(* IEC 61131-3 sources: 2026_Projet_YGO_ExcavatriceDragage/CODE_BACKUP/CODE_20260822_IntroductionTestCI/G_CYCLE, 6 files *)

(* ---- E_CycleStep.st ---- *)
(* =======================================================================
   ⚙️ E_CycleStep — Étapes de la machine d'état du cycle automatique
   ───────────────────────────────────────────────────────────────
   🎯 Rôle : Énumération des étapes du cycle automatique de dragage (X0 à X13 + STABILIZING)
   📄 Doc métier : DOC/AF/AF_Partie-04_Mode_SemiAuto_Sequenceur_v2.1.md
   ======================================================================= *)

TYPE E_CycleStep :
(
  X0_PREPARATION      := 0,   (* Début de graphe : à la TRÉMIE, treuils en position HAUTE *)
  X1_HOMING           := 1,   (* Vitesses lentes pour chercher capteur top + référencement *)
  X2_WORK_POS_SELECT  := 2,   (* Sélection cible Trémie/P1/Maintenance + translation validée *)
  X3_OPEN_BUCKET      := 3,   (* Ouverture benne (si déjà ouverte -> passe vite) *)
  X4_DESCEND_OPEN     := 4,   (* Plongée benne ouverte, M1+M2 synchro, Kobold mesure ON *)
  X5_BOTTOM_CONFIRMED := 5,   (* Fond validé (FB_DiveSearch) ; arrêt descente *)
  X6_CLOSE_BUCKET     := 6,   (* Fermeture benne — tolérance « à peu près fermé » *)
  X7_CTRL_ASCENT      := 7,   (* Remontée palier 1 de contrôle *)
  X8_ASCENT_LOADED    := 8,   (* Remontée nominale jusqu'à limite haute *)
  X9_DRAIN_PAUSE      := 9,   (* Égouttage temporisé — temps affiché IHM *)
  X10_TRANSLATE_DUMP  := 10,  (* Translation vers trémie + avertissements IHM *)
  X11_OPEN_DUMP       := 11,  (* Ouverture benne = vidage ; montée possible, descente ouvre *)
  X13_DONE_SYNC       := 13,  (* Fin de cycle, synchronisation finale (R4) + compteur *)
  STABILIZING         := 14   (* État d'attente/stabilisation — pas une erreur *)
);
END_TYPE

(* ---- E_DiveSearchState.st ---- *)
(* =======================================================================
   ⚙️ E_DiveSearchState — Phases internes de recherche du fond Kobold
   ───────────────────────────────────────────────────────────────
   🎯 Rôle : Énumération des phases de détection et recherche du fond
   📄 Doc métier : DOC/AF/AF_Partie-04_Mode_SemiAuto_Sequenceur_v2.1.md
   ======================================================================= *)

TYPE E_DiveSearchState :
(
    WAIT_PRECONDITIONS := 0, (* Attente benne ouverte, positions et Kobold au repos *)
    READY_TO_DESCEND   := 1, (* Prêt à assister une demande de descente *)
    SEARCHING_IMMERSION := 2, (* Descente : attente front 0->1 dans fenêtre eau *)
    SEARCHING_BOTTOM    := 3, (* Immersion validée : attente front 1->0 au fond *)
    BOTTOM_CONFIRMED    := 4, (* Fond validé ; extraction peut être demandée *)
    ERROR_HOLD          := 5  (* Séquence invalide, descente assistée interdite *)
);
END_TYPE

(* ---- E_ExtractionSequenceState.st ---- *)
(* =======================================================================
   ⚙️ E_ExtractionSequenceState — Phases d'extraction assistée
   ───────────────────────────────────────────────────────────────
   🎯 Rôle : Énumération des phases de la séquence d'extraction assistée
   📄 Doc métier : DOC/AF/AF_Partie-04_Mode_SemiAuto_Sequenceur_v2.1.md
   ======================================================================= *)

TYPE E_ExtractionSequenceState :
(
    WAIT_BOTTOM_CONFIRMATION := 0, (* Attente fond Kobold ou attestation opérateur *)
    READY_TO_CLOSE            := 1, (* Prêt à fermer la benne *)
    CLOSING_BUCKET            := 2, (* FB_Bucket ferme M2 seul *)
    CONTROL_ASCENT            := 3, (* M1/M2 synchronisés au palier sans contacteur vitesse *)
    NOMINAL_ASCENT            := 4, (* Montée couplée avec vitesse demandée opérateur *)
    ERROR_HOLD                := 5  (* Défaut extraction, reprise interdite avant reset *)
);
END_TYPE

(* ---- FB_Cycle.st ---- *)
(* =======================================================================
   ⚙️ FB_Cycle — Séquenceur du cycle automatique (Grafcet de dragage)
   ───────────────────────────────────────────────────────────────
   🎯 Rôle : Automate de cycle automatique de dragage (X0 à X13 + STABILIZING)
   🔒 Sécurité : Gating par mode et homme-mort, repli STABILIZING sur défaut
   🔌 Interface : Demandes de mouvements (treuils, translation, benne)
   📄 Doc métier : DOC/AF/AF_Partie-04_Mode_SemiAuto_Sequenceur_v2.1.md
   ======================================================================= *)

FUNCTION_BLOCK PUBLIC FB_Cycle
VAR_INPUT
    // === COMMANDES & AUTORISATIONS ===
    Enable                  : BOOL;         // --> [CMD] Activation generale du sequenceur
    Reset                   : BOOL;         // --> [CMD] Acquittement defaut (front)
    PowerContactorEngaged   : BOOL;         // --> [SAFE] Chaine de securite OK
    Mode                    : E_Mode;       // --> [CMD] Mode arbitre (SEMI_AUTO pour instance cycle)
    CycleMotionPermit       : BOOL;         // --> [CMD] Manche deflecte (non centre)
    DeadmanArmed            : BOOL;         // --> [CMD] Appui homme-mort (fenetre 3 s)
    HeartbeatIhmOk          : BOOL;         // --> [SAFE] IHM<->PLC valide

    // === COMMANDES OPERATEUR ===
    StartCycle              : BOOL;         // --> [CMD] Demande lancement / reprise (IHM)
    AbortCycle              : BOOL;         // --> [CMD] Demande abandon (IHM)

    // === CIBLES ET CONFIGURATION ===
    SelTarget               : INT;          // --> [CFG] Cible selectionnee (1=Tremie, 2=P2, 3=P1, 4=Maintenance)
    SetDepthM               : REAL;         // --> [CFG] Profondeur de consigne (negative)
    SetOffsetM              : REAL;         // --> [CFG] Ecart de fermeture benne cible

    // === FEEDBACKS CAPTEURS & MATERIEL ===
    KoboldContactFond       : BOOL;         // --> [HW] Retour dedie Kobold : TRUE = contact fond
    LimitLegalReached       : BOOL;         // --> [SAFE] Limite legale atteinte (descente interdite)
    LimitLegalDepthM        : REAL;         // --> [CFG] Profondeur legale minimale autorisee
    WinchSyncError          : BOOL;         // --> [SAFE] Desynchronisme bloquant M1/M2
    WinchSyncDeltaM         : REAL;         // --> [HW] Ecart codeurs M1/M2 pour diagnostic
    M1_CablePosM            : REAL;         // --> [HW] Position cable treuil M1 (recalee)
    M2_CablePosM            : REAL;         // --> [HW] Position cable treuil M2 (recalee)
    M1_MeasuredSpeedMps     : REAL;         // --> [HW] Vitesse lineaire mesuree M1 (m/s)
    M2_MeasuredSpeedMps     : REAL;         // --> [HW] Vitesse lineaire mesuree M2 (m/s)
    SpeedMismatchThresholdMps : REAL;       // --> [CFG] Seuil ecart vitesse ; 0 = controle desactive
    SpeedMismatchTimeout    : TIME;         // --> [CFG] Duree de confirmation ; 0 = controle desactive
    CableLimitM1AscentM     : REAL;         // --> [CFG] Limite haute d'exploitation M1

    // === FEEDBACKS TRANSLATION M3 ===
    Translation_At_P1           : BOOL;     // --> [HW] Capteur position P1 (arret travail)
    Translation_At_Tremie       : BOOL;     // --> [HW] Capteur fin de course tremie
    Translation_At_Maintenance : BOOL;     // --> [HW] Capteur fin de course maintenance
    Translation_Busy            : BOOL;     // --> [HW] Mouvement translation en cours
    Translation_Done            : BOOL;     // --> [HW] Cible translation atteinte

    // === FEEDBACKS BENNE ===
    Benne_Busy              : BOOL;         // --> [HW] Mouvement machoires benne en cours
    Benne_Done              : BOOL;         // --> [HW] Mouvement ouverture/fermeture termine
    Benne_IsOpen            : BOOL;         // --> [HW] Benne mecaniquement ouverte memorisee
    Benne_IsClosed          : BOOL;         // --> [HW] Benne mecaniquement fermee memorisee
    Benne_IsRoughlyClosed   : BOOL;         // --> [HW] Benne a peu pres fermee (tolerance matiere)

    // === REFERENCEMENT CODEURS ===
    HomedM1                 : BOOL;         // --> [HW] Codeur M1 reference
    HomedM2                 : BOOL;         // --> [HW] Codeur M2 reference
    TopPositionSensor       : BOOL;         // --> [HW] Capteur position haute (referencement)
    HomingRequest           : BOOL;         // --> [CMD] Demande de referencement (front)
END_VAR
VAR_OUTPUT
    // === ETATS IEC & DEFECTUOSITES ===
    Ready                   : BOOL;         // <-- [STAT] Sequenceur disponible
    Busy                    : BOOL;         // <-- [STAT] Cycle automatique actif
    Done                    : BOOL;         // <-- [STAT] Cycle automatique complete
    Error                   : BOOL;         // <-- [STAT] Defaut cycle
    ErrorId                 : WORD;         // <-- [DIAG] Code erreur bitmask
    SpeedMismatchMps        : REAL;         // <-- [DIAG] Ecart absolu vitesse M1/M2 (m/s)
    SpeedMismatchActive     : BOOL;         // <-- [DIAG] Seuil vitesse depasse sur cycle courant
    SpeedMismatchConfirmed  : BOOL;         // <-- [DIAG] Ecart vitesse confirme pendant timeout

    // === ORDRES ACTIONNEURS (COMMANDES STRUCTUREES) ===
    WinchM1Cmd              : ST_WinchCmdDemand;        // <-- [ACT] Demande treuil M1
    WinchM2Cmd              : ST_WinchCmdDemand;        // <-- [ACT] Demande treuil M2
    TranslationCmd          : ST_TranslationCmdDemand;  // <-- [ACT] Demande translation M3
    BucketCmd               : ST_BucketCmdDemand;       // <-- [ACT] Demande benne

    // === METADONNEES & SYNOPTIQUE ===
    CycleStep               : E_CycleStep;  // <-- [STAT] Etape active du Grafcet
    CycleStateStr           : STRING(80);   // <-- [STAT] Libelle en clair de l'etape
    CycleStepAtError        : E_CycleStep;  // <-- [DIAG] Etape specifique au moment du defaut
END_VAR
VAR_IN_OUT
    // === STRUCTURES PARTAGEES & COMPTEURS ===
    SampleCount             : INT;          // <-> [BUS] Compteur de prelevements (RETAIN)
END_VAR
VAR
    // === DETECTEURS DE FRONTS ===
    ResetEdge               : R_TRIG;       // . [LOC] Detecteur front montant Reset
    StartEdge               : R_TRIG;       // . [LOC] Detecteur front montant StartCycle
    DeadmanArmedEdge        : R_TRIG;       // . [LOC] Detecteur front montant DeadmanArmed (demarrage joystick)
    AbortEdge               : R_TRIG;       // . [LOC] Detecteur front montant AbortCycle
    ErrorEdge               : R_TRIG;       // . [LOC] Detecteur front montant Error

    // === ETATS INTERNES ===
    State                   : E_CycleStep := E_CycleStep.X0_PREPARATION; // . [LOC] Etape courante machine d'etat
    SavedState              : E_CycleStep := E_CycleStep.X0_PREPARATION; // . [LOC] Etape memorisee

    // === MEMORISATIONS & REGISTRES INTERNES ===
    TouchPositionM          : REAL;         // . [LOC] Position M1 memorisee lors du contact fond
    RaiseTargetM            : REAL;         // . [LOC] Profondeur de remontee memorisee
    SelectedWorkTarget      : INT;          // . [LOC] Cible de travail memorisee

    // === TEMPORISATEURS INTERNES ===
    DrainingTimer           : TON;          // . [LOC] Temporisateur de vidage (egouttage)
    StabilizationTimer      : TON;          // . [LOC] Temporisation maximale de remontee lente
    SpeedMismatchTimer      : TON;          // . [LOC] Confirmation temporelle ecart de vitesse
    StepMaxTimer            : TON;          // . [LOC] Tempo max d'etape

    // === CONSTANTES & CONFIGURATIONS INTERNES ===
    CtrlAscentDistM         : REAL := 2.0;      // . [LOC] Distance de remontee lente de controle
    CtrlAscentToleranceM    : REAL := 0.25;     // . [LOC] Ecart maximal admis entre codeurs
    CtrlAscentTimeout       : TIME := T#30s;    // . [LOC] Temps max pour zone de stabilisation
    DrainingTime            : TIME := T#5s;     // . [LOC] Temps d'egouttage par defaut
    StepMaxTimeout          : TIME := T#60s;    // . [LOC] Tempo max d'etape
END_VAR

// === IMPLEMENTATION ===

{region "§1 Gate securite"}
// 🛑 1. GATES DE SÉCURITÉ ET BLOCAGE (R8)
IF NOT Enable OR NOT PowerContactorEngaged THEN
    WinchM1Cmd.StartStop   := FALSE;
    WinchM1Cmd.Direction   := 0;
    WinchM1Cmd.SpeedPct    := 0.0;

    WinchM2Cmd.StartStop   := FALSE;
    WinchM2Cmd.Direction   := 0;
    WinchM2Cmd.SpeedPct    := 0.0;

    TranslationCmd.Start   := FALSE;
    TranslationCmd.Target  := 0;

    BucketCmd.Open         := FALSE;
    BucketCmd.Close        := FALSE;
    BucketCmd.KoboldContactorCmd := FALSE;

    State                := E_CycleStep.X0_PREPARATION;   // retour à la PREMIÈRE étape (R8)
    CycleStep            := E_CycleStep.X0_PREPARATION;
    CycleStateStr        := 'X0 - Désactivé : sécurité absente ou auto désactivé';
    Ready                := FALSE;
    Busy                 := FALSE;
    Done                 := FALSE;
    RETURN;
END_IF;
{endregion}

{region "§2 Preparation surveillance et commandes cycle"}
Ready := TRUE;
ResetEdge(CLK := Reset);
StartEdge(CLK := StartCycle);
DeadmanArmedEdge(CLK := DeadmanArmed);
AbortEdge(CLK := AbortCycle);
ErrorEdge(CLK := Error);

// 🧊 R9 — capture l'étape spécifique AVANT la bascule vers STABILIZING
IF ErrorEdge.Q THEN
    CycleStepAtError := State;
END_IF;

// ⏱️ Surveillance indépendante de la remontée lente
StabilizationTimer(IN := (State = E_CycleStep.X7_CTRL_ASCENT), PT := CtrlAscentTimeout);

// 📏 Comparaison vitesse réelle M1/M2
SpeedMismatchMps := ABS(M1_MeasuredSpeedMps - M2_MeasuredSpeedMps);
SpeedMismatchActive := (State = E_CycleStep.X7_CTRL_ASCENT)
                       AND CycleMotionPermit
                       AND (SpeedMismatchThresholdMps > 0.0)
                       AND (SpeedMismatchTimeout > T#0ms)
                       AND (SpeedMismatchMps > SpeedMismatchThresholdMps);
SpeedMismatchTimer(IN := SpeedMismatchActive, PT := SpeedMismatchTimeout);
SpeedMismatchConfirmed := SpeedMismatchTimer.Q;

// Tempo max d'étape (R5) — lancée SEULEMENT si pilotage joystick actif (pas de défaut au repos)
StepMaxTimer(IN := CycleMotionPermit AND (State <> E_CycleStep.X0_PREPARATION)
                  AND (State <> E_CycleStep.X13_DONE_SYNC)
                  AND (State <> E_CycleStep.STABILIZING),
             PT := StepMaxTimeout);

IF ResetEdge.Q THEN
    Error := FALSE;
    ErrorId := 16#0000;
    SavedState := E_CycleStep.X0_PREPARATION;
    IF State = E_CycleStep.STABILIZING THEN
        State := E_CycleStep.X0_PREPARATION;
    END_IF;
END_IF;

// 💓 Perte IHM : repli mémorisé. La reconnexion seule ne relance jamais le cycle.
IF NOT HeartbeatIhmOk AND State <> E_CycleStep.STABILIZING THEN
    Error := TRUE;
    ErrorId := ErrorId OR 16#0020;
    State := E_CycleStep.STABILIZING;
END_IF;

// Défaut de synchronisme : arrêt sûr et acquittement obligatoire.
IF WinchSyncError AND State <> E_CycleStep.STABILIZING THEN
    Error := TRUE;
    ErrorId := ErrorId OR 16#0002;
    State := E_CycleStep.STABILIZING;
END_IF;

// 🛡️ Écart de vitesse confirmé : arrêt du cycle et STABILIZING.
IF SpeedMismatchConfirmed AND State <> E_CycleStep.STABILIZING THEN
    Error := TRUE;
    ErrorId := ErrorId OR 16#0010;
    State := E_CycleStep.STABILIZING;
END_IF;

// Tempo max d'étape dépassée (blocage probable) → défaut
IF StepMaxTimer.Q AND State <> E_CycleStep.STABILIZING THEN
    Error := TRUE;
    ErrorId := ErrorId OR 16#0040;
    State := E_CycleStep.STABILIZING;
END_IF;

// Gestion de l'Abandon (D3 — pas de Pause)
IF AbortEdge.Q THEN
    State := E_CycleStep.X0_PREPARATION;
END_IF;
{endregion}

{region "§3 Machine etat cycle automatique"}
// 🔁 2. LOGIQUE DU SÉQUENCEUR (Machine d'état) — CASE sur enum unique (R1)
CASE State OF

    E_CycleStep.X0_PREPARATION:
        CycleStep := E_CycleStep.X0_PREPARATION;
        CycleStateStr := 'X0 - Vérification cohérence système';
        WinchM1Cmd.StartStop := FALSE; WinchM1Cmd.Direction := 0; WinchM1Cmd.SpeedPct := 0.0;
        WinchM2Cmd.StartStop := FALSE; WinchM2Cmd.Direction := 0; WinchM2Cmd.SpeedPct := 0.0;
        TranslationCmd.Start := FALSE; TranslationCmd.Target := 0;
        BucketCmd.Open := FALSE; BucketCmd.Close := FALSE; BucketCmd.KoboldContactorCmd := FALSE;
        Busy := FALSE; Done := FALSE;

        // Transition si système sain et réarmé (front reset ou démarrage).
        // 🔫 D2 : démarrage par bouton IHM (StartEdge) OU armement homme-mort joystick
        // (DeadmanArmedEdge) — l'opérateur peut lancer depuis l'IHM ou le joystick.
        // La continuité des mouvements ne dépend que de CycleMotionPermit (manche défléchi).
        IF StartEdge.Q OR DeadmanArmedEdge.Q THEN
            State := E_CycleStep.X1_HOMING;
        END_IF;

    E_CycleStep.X1_HOMING:
        CycleStep := E_CycleStep.X1_HOMING;
        CycleStateStr := 'X1 - Référencement codeurs (vitesses lentes)';
        Busy := TRUE;

        // Vitesses lentes pour chercher capteur top + référencement
        IF NOT HomedM1 OR NOT HomedM2 THEN
            WinchM1Cmd.StartStop := CycleMotionPermit;
            WinchM1Cmd.Direction := 1;   // montée lente vers capteur top
            WinchM1Cmd.SpeedPct := 10.0;
            WinchM2Cmd.StartStop := CycleMotionPermit;
            WinchM2Cmd.Direction := 1;
            WinchM2Cmd.SpeedPct := 10.0;
            IF HomingRequest THEN
                // déclenche le référencement (via FB_Encoder_Homing en aval)
                State := E_CycleStep.X2_WORK_POS_SELECT;
            END_IF;
        ELSE
            // déjà homé → passe vite
            State := E_CycleStep.X2_WORK_POS_SELECT;
        END_IF;

    E_CycleStep.X2_WORK_POS_SELECT:
        CycleStep := E_CycleStep.X2_WORK_POS_SELECT;
        CycleStateStr := 'X2 - Sélection position travail';
        Busy := TRUE;

        // Destinations sélectionnables : Trémie(1), P1(3), Maintenance(4).
        // P2(2) n'est PAS une destination — capteur de passage en petite vitesse (PV).
        // Si aucune cible valide n'est sélectionnée, on ATTEND à X2 (pas de défaut) :
        // l'opérateur choisit la position de travail via l'IHM (SelTarget).
        IF (SelTarget = 1) OR (SelTarget = 3) OR (SelTarget = 4) THEN
            SelectedWorkTarget := SelTarget;
            TranslationCmd.Target := SelTarget;
            TranslationCmd.Start := CycleMotionPermit;
            // Arrivée à la cible (Trémie/P1/Maintenance) — capteurs PV/PVP2/P2 = ralentissement
            IF CycleMotionPermit AND (
                (SelTarget = 1 AND Translation_At_Tremie) OR
                (SelTarget = 3 AND Translation_At_P1) OR
                (SelTarget = 4 AND Translation_At_Maintenance)) THEN
                TranslationCmd.Start := FALSE;
                State := E_CycleStep.X3_OPEN_BUCKET;
            END_IF;
        END_IF;

    E_CycleStep.X3_OPEN_BUCKET:
        CycleStep := E_CycleStep.X3_OPEN_BUCKET;
        CycleStateStr := 'X3 - Ouverture benne';
        Busy := TRUE;

        // Ouverture benne ; si déjà ouverte → passe vite
        IF Benne_IsOpen THEN
            State := E_CycleStep.X4_DESCEND_OPEN;
        ELSE
            BucketCmd.Open := CycleMotionPermit;
            IF CycleMotionPermit AND Benne_Done AND Benne_IsOpen THEN
                BucketCmd.Open := FALSE;
                State := E_CycleStep.X4_DESCEND_OPEN;
            END_IF;
        END_IF;

    E_CycleStep.X4_DESCEND_OPEN:
        CycleStep := E_CycleStep.X4_DESCEND_OPEN;
        CycleStateStr := 'X4 - Plongée benne ouverte (synchro)';

        // M1 et M2 descendent ensemble (synchro gérée en aval)
        WinchM1Cmd.StartStop := CycleMotionPermit;
        WinchM1Cmd.Direction := -1;
        WinchM1Cmd.SpeedPct  := 50.0;
        WinchM2Cmd.StartStop := CycleMotionPermit;
        WinchM2Cmd.Direction := -1;
        WinchM2Cmd.SpeedPct  := 50.0;
        BucketCmd.KoboldContactorCmd := TRUE;

        // Transition uniquement sur le retour dédié Kobold.
        IF CycleMotionPermit AND KoboldContactFond THEN
            WinchM1Cmd.StartStop := FALSE;
            WinchM2Cmd.StartStop := FALSE;
            BucketCmd.KoboldContactorCmd := FALSE;
            TouchPositionM := M1_CablePosM;
            IF LimitLegalDepthM < -0.01 THEN
                RaiseTargetM := MAX(TouchPositionM + 0.5, LimitLegalDepthM + 0.5);
            ELSE
                RaiseTargetM := TouchPositionM + 0.5;
            END_IF;
            State := E_CycleStep.X5_BOTTOM_CONFIRMED;
        ELSIF LimitLegalReached THEN
            Error := TRUE;
            ErrorId := ErrorId OR 16#0001;
            WinchM1Cmd.StartStop := FALSE;
            WinchM2Cmd.StartStop := FALSE;
            BucketCmd.KoboldContactorCmd := FALSE;
            State := E_CycleStep.STABILIZING;
        END_IF;

    E_CycleStep.X5_BOTTOM_CONFIRMED:
        CycleStep := E_CycleStep.X5_BOTTOM_CONFIRMED;
        CycleStateStr := 'X5 - Fond confirmé : remontée sécurisée';

        WinchM1Cmd.StartStop := CycleMotionPermit;
        WinchM1Cmd.Direction := 1;
        WinchM1Cmd.SpeedPct := 20.0;
        WinchM2Cmd.StartStop := CycleMotionPermit;
        WinchM2Cmd.Direction := 1;
        WinchM2Cmd.SpeedPct := 20.0;

        // Les deux treuils restent synchronisés jusqu'au-dessus de la limite légale.
        IF CycleMotionPermit AND (M1_CablePosM >= RaiseTargetM) AND (M2_CablePosM >= RaiseTargetM) THEN
            WinchM1Cmd.StartStop := FALSE;
            WinchM2Cmd.StartStop := FALSE;
            State := E_CycleStep.X6_CLOSE_BUCKET;
        END_IF;

    E_CycleStep.X6_CLOSE_BUCKET:
        CycleStep := E_CycleStep.X6_CLOSE_BUCKET;
        CycleStateStr := 'X6 - Fermeture benne (tolérance à peu près fermé)';

        WinchM1Cmd.StartStop := FALSE;
        BucketCmd.Close := TRUE;

        // Tolérance : si benne « à peu près fermée » (matière/objet), on remonte et on contrôle
        IF CycleMotionPermit AND (Benne_Done AND (Benne_IsClosed OR Benne_IsRoughlyClosed)) THEN
            BucketCmd.Close := FALSE;
            State := E_CycleStep.X7_CTRL_ASCENT;
        END_IF;

    E_CycleStep.X7_CTRL_ASCENT:
        CycleStep := E_CycleStep.X7_CTRL_ASCENT;
        CycleStateStr := 'X7 - Remontée lente de contrôle';

        WinchM1Cmd.StartStop := CycleMotionPermit;
        WinchM1Cmd.Direction := 1;
        WinchM1Cmd.SpeedPct  := 20.0;
        WinchM2Cmd.StartStop := CycleMotionPermit;
        WinchM2Cmd.Direction := 1;
        WinchM2Cmd.SpeedPct  := 20.0;

        // Contrôle des deux codeurs
        IF WinchSyncError OR (ABS(M1_CablePosM - M2_CablePosM) > CtrlAscentToleranceM) THEN
            Error := TRUE;
            ErrorId := ErrorId OR 16#0008;
            State := E_CycleStep.STABILIZING;
        ELSIF CycleMotionPermit
           AND (M1_CablePosM >= (TouchPositionM + CtrlAscentDistM))
           AND (M2_CablePosM >= (TouchPositionM + CtrlAscentDistM))
           AND (ABS(M1_CablePosM - M2_CablePosM) <= CtrlAscentToleranceM) THEN
            State := E_CycleStep.X8_ASCENT_LOADED;
        ELSIF StabilizationTimer.Q THEN
            Error := TRUE;
            ErrorId := ErrorId OR 16#0008;
            State := E_CycleStep.STABILIZING;
        END_IF;

    E_CycleStep.X8_ASCENT_LOADED:
        CycleStep := E_CycleStep.X8_ASCENT_LOADED;
        CycleStateStr := 'X8 - Remontée en charge';

        WinchM1Cmd.StartStop := CycleMotionPermit;
        WinchM1Cmd.Direction := 1;
        WinchM1Cmd.SpeedPct  := 70.0;
        WinchM2Cmd.StartStop := CycleMotionPermit;
        WinchM2Cmd.Direction := 1;
        WinchM2Cmd.SpeedPct  := 70.0;

        // Transition alignée sur la limite haute d'exploitation
        IF CycleMotionPermit AND M1_CablePosM >= CableLimitM1AscentM THEN
            WinchM1Cmd.StartStop := FALSE;
            WinchM2Cmd.StartStop := FALSE;
            State := E_CycleStep.X9_DRAIN_PAUSE;
        END_IF;

    E_CycleStep.X9_DRAIN_PAUSE:
        CycleStep := E_CycleStep.X9_DRAIN_PAUSE;
        CycleStateStr := 'X9 - Égouttage du godet en cours';
        WinchM1Cmd.StartStop := FALSE;
        WinchM2Cmd.StartStop := FALSE;

        DrainingTimer(IN := TRUE, PT := DrainingTime);
        // Temps écoulé affiché IHM (CycleStateStr + champ dédié)
        IF CycleMotionPermit AND DrainingTimer.Q THEN
            DrainingTimer(IN := FALSE);
            State := E_CycleStep.X10_TRANSLATE_DUMP;
        END_IF;

    E_CycleStep.X10_TRANSLATE_DUMP:
        CycleStep := E_CycleStep.X10_TRANSLATE_DUMP;
        CycleStateStr := 'X10 - Déplacement vers trémie (grille/crible libres)';

        TranslationCmd.Target := 1; // Trémie
        TranslationCmd.Start := CycleMotionPermit;

        // Avertissement IHM : grille abaissée/libre, crible libre pour réceptionner la charge
        // (porté par CycleStateStr + OperatorAction côté supervision)

        // Transition si translation arrivé à la trémie
        IF CycleMotionPermit AND Translation_At_Tremie THEN
            TranslationCmd.Start := FALSE;
            State := E_CycleStep.X11_OPEN_DUMP;
        END_IF;

    E_CycleStep.X11_OPEN_DUMP:
        CycleStep := E_CycleStep.X11_OPEN_DUMP;
        CycleStateStr := 'X11 - Vidange / ouverture du godet (montée possible, descente ouvre)';

        // Montée possible (treuils vers le haut) ; descente fait ouvrir la benne.
        // Montée : on laisse l'opérateur remonter les 2 treuils en synchro si besoin.
        WinchM1Cmd.StartStop := CycleMotionPermit AND (WinchM1Cmd.Direction = 1);
        WinchM1Cmd.Direction := 1;
        WinchM1Cmd.SpeedPct  := 20.0;
        WinchM2Cmd.StartStop := CycleMotionPermit AND (WinchM2Cmd.Direction = 1);
        WinchM2Cmd.Direction := 1;
        WinchM2Cmd.SpeedPct  := 20.0;

        // Descente → ouverture benne (vidage)
        BucketCmd.Open := CycleMotionPermit AND (WinchM1Cmd.Direction = -1);

        // Contrôle convoyeurs par MESSAGE utilisateur (pas encore câblé) :
        // CycleStateStr + OperatorAction côté supervision demandent de vérifier
        // que les convoyeurs sont en route avant/au lâcher.
        IF CycleMotionPermit AND Benne_Done AND Benne_IsOpen THEN
            BucketCmd.Open := FALSE;
            State := E_CycleStep.X13_DONE_SYNC;
        END_IF;

    E_CycleStep.X13_DONE_SYNC:
        CycleStep := E_CycleStep.X13_DONE_SYNC;
        CycleStateStr := 'X13 - Cycle automatique complété - prêt';
        WinchM1Cmd.StartStop := FALSE;
        WinchM2Cmd.StartStop := FALSE;
        TranslationCmd.Start := FALSE;
        Done := TRUE;
        Busy := FALSE;

        // Compteur de prélèvements (RETAIN, Q3bis) — compte inconditionnellement
        SampleCount := SampleCount + 1;

        // Rebouclage sur X0_PREPARATION (trémie, treuils hauts) — pas de retour P1
        IF StartEdge.Q THEN
            Done := FALSE;
            State := E_CycleStep.X0_PREPARATION;
        END_IF;

    E_CycleStep.STABILIZING:
        CycleStep := E_CycleStep.STABILIZING;
        CycleStateStr := 'X14 - Cycle en attente / stabilisation (STAB)';
        WinchM1Cmd.StartStop := FALSE;
        WinchM2Cmd.StartStop := FALSE;
        TranslationCmd.Start := FALSE;
        BucketCmd.Open := FALSE;
        BucketCmd.Close := FALSE;

END_CASE;
{endregion}

{region "§4 Repli homme mort"}
// 🛑 Relâchement du manche (retour au centre) : aucune demande d'actionneur ne reste active.
// L'étape est mémorisée et reprend au prochain appui valide (D2).
IF Busy AND NOT CycleMotionPermit THEN
    WinchM1Cmd.StartStop := FALSE;
    WinchM2Cmd.StartStop := FALSE;
    TranslationCmd.Start := FALSE;
    BucketCmd.Open := FALSE;
    BucketCmd.Close := FALSE;
    BucketCmd.KoboldContactorCmd := FALSE;
END_IF;
{endregion}

END_FUNCTION_BLOCK

(* ---- FB_DiveSearch.st ---- *)
(* =======================================================================
   ⚙️ FB_DiveSearch — Assistance plongée et recherche du fond Kobold
   ───────────────────────────────────────────────────────────────
   🎯 Rôle : Qualification du capteur Kobold et autorisation de descente
   🛡️ Sécurité : Verrouillage si séquence d'immersion 0->1->0 invalide
   🔌 Interface : Intention de descente et mesures vers permis de descente
   📄 Doc métier : DOC/AF/AF_Partie-04_Mode_SemiAuto_Sequenceur_v2.1.md
   ======================================================================= *)
FUNCTION_BLOCK FB_DiveSearch
VAR_INPUT
    // === COMMANDES & AUTORISATIONS ===
    Enable                  : BOOL;         // --> [CMD] Activation generale du FB (TRUE=Autorise)
    Reset                   : BOOL;         // --> [CMD] Acquittement defaut (front)
    PowerContactorEngaged   : BOOL;         // --> [SAFE] Chaine de securite OK
    Mode                    : E_Mode;       // --> [CMD] Mode de fonctionnement arbitre
    MotionRequestActive     : BOOL;         // --> [CMD] Intention de mouvement active
    MotionDirection         : INT;          // --> [CMD] Sens de mouvement (-1 = descente)

    // === CAPTEURS & ETATS BENNE ===
    BucketIsOpen            : BOOL;         // --> [HW] Benne ouverte confirmee
    KoboldImmersed          : BOOL;         // --> [HW] Capteur Kobold immerge (FALSE=hors eau, TRUE=immerge)
    M1Position_M            : REAL;         // --> [HW] Position codeur treuil M1 (m)
    M2Position_M            : REAL;         // --> [HW] Position codeur treuil M2 (m)
    PositionsValid          : BOOL;         // --> [HW] Validite des mesures de position

    // === CONFIGURATION & SEUILS ===
    DiveStartMin_M          : REAL;         // --> [CFG] Seuil position min pour debut plongee (m)
    ImmersionUpper_M        : REAL;         // --> [CFG] Borne haute fenetre d'immersion (m)
    ImmersionLower_M        : REAL;         // --> [CFG] Borne basse fenetre d'immersion (m)
    BypassPreconditions     : BOOL := FALSE;// --> [TST] Bypass preconditions et seuils (mode test)
END_VAR
VAR_OUTPUT
    // === ETATS IEC & DEFECTUOSITES ===
    Ready                   : BOOL;         // <-- [STAT] FB pret a fonctionner
    // Status.ErrorId : bit0 precond, bit1 seq, bit2 cfg
    Status                  : ST_FbStatus;  // <-- [STAT] Etat global FB (Busy/Done/Error/ErrorId/State/StateAtError)
    DiveState               : E_DiveSearchState; // <-- [STAT] Phase interne de recherche fond

    // === PERMIS & AUTORISATIONS ===
    DescendPermit           : BOOL;         // <-- [ACT] Autorisation de descente assistee
    KoboldMeasureEnable     : BOOL;         // <-- [ACT] Activation mesure/acquisition Kobold
    BottomTouchConfirmed    : BOOL;         // <-- [STAT] Contact fond valide et confirme

    // === DIAGNOSTIC IHM ===
    OperatorActionId        : WORD;         // <-- [DIAG] ID action operateur requise
    OperatorAction          : STRING(120);  // <-- [DIAG] Message explicatif operateur
END_VAR
VAR
    // === DETECTEURS DE FRONTS ===
    ResetEdge               : R_TRIG;       // . [LOC] Detecteur front montant Reset
    KoboldRiseEdge          : R_TRIG;       // . [LOC] Detecteur front entrant eau (0->1)
    KoboldFallEdge          : F_TRIG;       // . [LOC] Detecteur front sortie eau / fond (1->0)

    // === VARIABLES LOCALES INTERNES ===
    ImmersionConfirmed      : BOOL;         // . [LOC] Immersion dans la fenetre d'eau validee
    ErrorCausePresent       : BOOL;         // . [LOC] Presence d'une cause de defaut parametrage
END_VAR

{region "§1 Gate desactivation"}
IF NOT Enable OR NOT PowerContactorEngaged THEN
    Ready := FALSE; Status.Busy := FALSE; Status.Done := FALSE;
    DescendPermit := FALSE; KoboldMeasureEnable := FALSE;
    BottomTouchConfirmed := FALSE;
    Status.State := E_State.DISABLED;
    Status.StateAtError := E_State.DISABLED;
    DiveState := E_DiveSearchState.WAIT_PRECONDITIONS;
    OperatorActionId := 0; OperatorAction := '';
    ImmersionConfirmed := FALSE;
    RETURN;
END_IF;

{endregion}

{region "§2 Preconditions fronts et rearmement"}
ResetEdge(CLK := Reset);
KoboldRiseEdge(CLK := KoboldImmersed);
KoboldFallEdge(CLK := KoboldImmersed);

ErrorCausePresent := NOT BypassPreconditions AND ((DiveStartMin_M < ImmersionUpper_M)
                  OR (ImmersionUpper_M <= ImmersionLower_M));
IF ErrorCausePresent THEN
    Status.ErrorId := Status.ErrorId OR 16#0004;
END_IF;

(* Reset = front + causes disparues ; aucun redémarrage automatique. *)
IF ResetEdge.Q AND NOT ErrorCausePresent AND NOT KoboldImmersed AND NOT MotionRequestActive THEN
    Status.ErrorId := 16#0000;
    ImmersionConfirmed := FALSE;
    BottomTouchConfirmed := FALSE;
    Status.StateAtError := E_State.DISABLED;
    DiveState := E_DiveSearchState.WAIT_PRECONDITIONS;
END_IF;

DescendPermit := FALSE; KoboldMeasureEnable := FALSE;
Ready := FALSE; Status.Busy := FALSE; Status.Done := FALSE;
OperatorActionId := 0; OperatorAction := '';

{endregion}

{region "§3 Machine etat plongee recherche fond"}
IF Status.ErrorId <> 16#0000 THEN
    Status.State := E_State.READY;
    DiveState := E_DiveSearchState.ERROR_HOLD;
    OperatorActionId := 16#0180;
    OperatorAction := 'Vérifier les conditions puis réarmer avant une nouvelle plongée.';
ELSE
    CASE DiveState OF
        E_DiveSearchState.WAIT_PRECONDITIONS:
            Status.State := E_State.INIT;
            IF NOT BypassPreconditions
               AND (NOT BucketIsOpen OR NOT PositionsValid OR KoboldImmersed
                    OR (M1Position_M < DiveStartMin_M) OR (M2Position_M < DiveStartMin_M)) THEN
                OperatorActionId := 16#0100;
                OperatorAction := 'Vérifier les conditions initiales de plongée.';
            ELSE
                DiveState := E_DiveSearchState.READY_TO_DESCEND;
            END_IF;

        E_DiveSearchState.READY_TO_DESCEND:
            Status.State := E_State.READY;
            Ready := TRUE;
            OperatorActionId := 16#0101;
            OperatorAction := 'Demander une descente pour rechercher le fond.';
            IF MotionRequestActive AND (MotionDirection = -1) THEN
                DiveState := E_DiveSearchState.SEARCHING_IMMERSION;
            END_IF;

        E_DiveSearchState.SEARCHING_IMMERSION:
            Status.State := E_State.BUSY;
            Status.Busy := TRUE;
            DescendPermit := MotionRequestActive AND (MotionDirection = -1);
            KoboldMeasureEnable := TRUE;
            OperatorActionId := 16#0102;
            OperatorAction := 'Maintenir la descente : recherche immersion Kobold.';
            IF KoboldRiseEdge.Q THEN
                IF (M1Position_M <= ImmersionUpper_M) AND (M1Position_M >= ImmersionLower_M)
                   AND (M2Position_M <= ImmersionUpper_M) AND (M2Position_M >= ImmersionLower_M) THEN
                    ImmersionConfirmed := TRUE;
                    DiveState := E_DiveSearchState.SEARCHING_BOTTOM;
                ELSE
                    Status.ErrorId := Status.ErrorId OR 16#0002;
                    Status.StateAtError := Status.State;
                END_IF;
            ELSIF (M1Position_M < ImmersionLower_M) OR (M2Position_M < ImmersionLower_M) THEN
                Status.ErrorId := Status.ErrorId OR 16#0002;
                Status.StateAtError := Status.State;
            END_IF;

        E_DiveSearchState.SEARCHING_BOTTOM:
            Status.State := E_State.BUSY;
            Status.Busy := TRUE;
            DescendPermit := MotionRequestActive AND (MotionDirection = -1);
            KoboldMeasureEnable := TRUE;
            OperatorActionId := 16#0103;
            OperatorAction := 'Maintenir la descente : immersion validée, recherche du fond.';
            IF KoboldFallEdge.Q AND ImmersionConfirmed THEN
                BottomTouchConfirmed := TRUE;
                ImmersionConfirmed := FALSE;
                DiveState := E_DiveSearchState.BOTTOM_CONFIRMED;
            END_IF;

        E_DiveSearchState.BOTTOM_CONFIRMED:
            Status.State := E_State.DONE;
            Status.Done := TRUE;
            OperatorActionId := 16#0104;
            OperatorAction := 'Fond détecté : demander la fermeture ou l extraction.';

        E_DiveSearchState.ERROR_HOLD:
            Status.State := E_State.READY;
    END_CASE;
END_IF;

Status.Error := (Status.ErrorId <> 16#0000);

{endregion}

(* ---- FB_ExtractionSequence.st ---- *)
(* =======================================================================
   ⚙️ FB_ExtractionSequence — Fermeture benne et remontée assistée
   ───────────────────────────────────────────────────────────────
   🎯 Rôle : Séquence d'extraction (fermeture benne, remontée de contrôle, remontée nominale)
   🛡️ Sécurité : Aucune remontée assistée sans fond confirmé, contrôle palier 1
   📄 Doc métier : DOC/AF/AF_Partie-04_Mode_SemiAuto_Sequenceur_v2.1.md
   ======================================================================= *)
FUNCTION_BLOCK FB_ExtractionSequence
VAR_INPUT
    // === COMMANDES & AUTORISATIONS ===
    Enable                      : BOOL;     // --> [CMD] Activation generale du FB (TRUE=Autorise)
    Reset                       : BOOL;     // --> [CMD] Acquittement defaut (front)
    PowerContactorEngaged       : BOOL;     // --> [SAFE] Chaine de securite OK
    Mode                        : E_Mode;   // --> [CMD] Mode de fonctionnement arbitre
    MotionRequestActive         : BOOL;     // --> [CMD] Intention de mouvement active
    MotionDirection             : INT;      // --> [CMD] Sens de mouvement (+1 = montee)
    BottomPositionConfirmed     : BOOL;     // --> [SAFE] Attestation fond confirme (Kobold ou op)

    // === CAPTEURS & ETATS MATERIELS ===
    BucketIsClosed              : BOOL;     // --> [HW] Benne fermee confirmee
    BucketBusy                  : BOOL;     // --> [HW] Mouvement benne en cours
    BucketError                 : BOOL;     // --> [SAFE] Defaut sur sous-systeme benne
    WinchSyncError              : BOOL;     // --> [SAFE] Defaut de desynchronisme treuils M1/M2
    M1Position_M                : REAL;     // --> [HW] Position codeur treuil M1 (m)
    M2Position_M                : REAL;     // --> [HW] Position codeur treuil M2 (m)
    M1MeasuredSpeedValid        : BOOL;     // --> [HW] Validite mesure vitesse M1
    M2MeasuredSpeedValid        : BOOL;     // --> [HW] Validite mesure vitesse M2
    PositionsValid              : BOOL;     // --> [HW] Validite des mesures de position

    // === CONFIGURATION & REGLAGES ===
    ControlAscentDistance_M     : REAL;     // --> [CFG] Distance palier 1 de controle remontee (m)
END_VAR
VAR_OUTPUT
    // === ETATS IEC & DEFECTUOSITES ===
    Ready                       : BOOL;     // <-- [STAT] FB pret a fonctionner (sortie libre, hors ST_FbStatus)
    // 🧩 Statut transverse (forme cible) — regroupe Busy/Done/Error/ErrorId/State/StateAtError.
    // ErrorId bit0:fond ; bit1:ferme ; bit2:ctrl ; bit3:cfg.
    Status                      : ST_FbStatus; // <-- [STAT] Etat global FB (Busy/Done/Error/ErrorId/State/StateAtError)
    ExtractionState             : E_ExtractionSequenceState; // <-- [STAT] Phase interne extraction

    // === ORDRES & AUTORISATIONS ===
    BucketCloseRequest          : BOOL;     // <-- [ACT] Demande de fermeture benne
    AscentPermit                : BOOL;     // <-- [ACT] Autorisation de remontee assistee
    ForceMinSpeedStep           : BOOL;     // <-- [ACT] Forcage vitesse minimale (palier de controle)
    BottomConfirmationConsumed  : BOOL;     // <-- [STAT] Signal confirmation fond consomme

    // === DIAGNOSTIC IHM ===
    OperatorActionId            : WORD;     // <-- [DIAG] ID action operateur requise
    OperatorAction              : STRING(120); // <-- [DIAG] Message explicatif operateur
END_VAR
VAR
    // === DETECTEURS DE FRONTS ===
    ResetEdge                   : R_TRIG;   // . [LOC] Detecteur front montant Reset

    // === MEMORISATIONS & POSITIONS INTERNES ===
    ControlStartM1Position_M    : REAL;     // . [LOC] Position M1 au debut du palier de controle (m)
    ControlStartM2Position_M    : REAL;     // . [LOC] Position M2 au debut du palier de controle (m)

    // === VARIABLES LOCALES INTERNES ===
    ErrorCausePresent           : BOOL;     // . [LOC] Presence d'une cause de defaut parametrage
END_VAR

{region "§1 Gate desactivation"}
IF NOT Enable OR NOT PowerContactorEngaged THEN
    Ready := FALSE; Status.Busy := FALSE; Status.Done := FALSE;
    BucketCloseRequest := FALSE; AscentPermit := FALSE; ForceMinSpeedStep := FALSE;
    BottomConfirmationConsumed := FALSE;
    Status.State := E_State.DISABLED;
    Status.StateAtError := E_State.DISABLED;
    ExtractionState := E_ExtractionSequenceState.WAIT_BOTTOM_CONFIRMATION;
    OperatorActionId := 0; OperatorAction := '';
    RETURN;
END_IF;

{endregion}

{region "§2 Preconditions reset et initialisation sorties"}
ResetEdge(CLK := Reset);
ErrorCausePresent := (ControlAscentDistance_M <= 0.0);
IF ErrorCausePresent THEN
    Status.ErrorId := Status.ErrorId OR 16#0008;
END_IF;
IF ResetEdge.Q AND NOT ErrorCausePresent AND NOT MotionRequestActive THEN
    Status.ErrorId := 16#0000;
    Status.StateAtError := E_State.DISABLED;
    ExtractionState := E_ExtractionSequenceState.WAIT_BOTTOM_CONFIRMATION;
END_IF;

Ready := FALSE; Status.Busy := FALSE; Status.Done := FALSE;
BucketCloseRequest := FALSE; AscentPermit := FALSE; ForceMinSpeedStep := FALSE;
BottomConfirmationConsumed := FALSE;
OperatorActionId := 0; OperatorAction := '';

{endregion}

{region "§3 Machine etat fermeture remontee"}
IF Status.ErrorId <> 16#0000 THEN
    Status.State := E_State.READY;
    ExtractionState := E_ExtractionSequenceState.ERROR_HOLD;
    OperatorActionId := 16#0280;
    OperatorAction := 'Vérifier la benne et les treuils puis réarmer avant de reprendre.';
ELSE
    CASE ExtractionState OF
        E_ExtractionSequenceState.WAIT_BOTTOM_CONFIRMATION:
            Status.State := E_State.INIT;
            IF BottomPositionConfirmed THEN
                ExtractionState := E_ExtractionSequenceState.READY_TO_CLOSE;
            ELSE
                OperatorActionId := 16#0200;
                OperatorAction := 'Confirmer que la benne est posée au fond avant extraction.';
            END_IF;

        E_ExtractionSequenceState.READY_TO_CLOSE:
            Status.State := E_State.READY;
            Ready := TRUE;
            OperatorActionId := 16#0201;
            OperatorAction := 'Demander la montée pour fermer la benne.';
            IF MotionRequestActive AND (MotionDirection = 1) THEN
                BottomConfirmationConsumed := TRUE;
                ExtractionState := E_ExtractionSequenceState.CLOSING_BUCKET;
            END_IF;

        E_ExtractionSequenceState.CLOSING_BUCKET:
            Status.State := E_State.BUSY;
            Status.Busy := TRUE;
            BucketCloseRequest := MotionRequestActive AND (MotionDirection = 1);
            OperatorActionId := 16#0202;
            OperatorAction := 'Maintenir la montée : fermeture de la benne en cours.';
            IF BucketError THEN
                Status.ErrorId := Status.ErrorId OR 16#0002;
                Status.StateAtError := Status.State;
            ELSIF BucketIsClosed AND NOT BucketBusy THEN
                ControlStartM1Position_M := M1Position_M;
                ControlStartM2Position_M := M2Position_M;
                ExtractionState := E_ExtractionSequenceState.CONTROL_ASCENT;
            END_IF;

        E_ExtractionSequenceState.CONTROL_ASCENT:
            Status.State := E_State.BUSY;
            Status.Busy := TRUE;
            AscentPermit := MotionRequestActive AND (MotionDirection = 1);
            ForceMinSpeedStep := TRUE;
            OperatorActionId := 16#0203;
            OperatorAction := 'Maintenir la montée : contrôle charge au palier minimal.';
            IF WinchSyncError OR NOT PositionsValid OR NOT M1MeasuredSpeedValid OR NOT M2MeasuredSpeedValid THEN
                Status.ErrorId := Status.ErrorId OR 16#0004;
                Status.StateAtError := Status.State;
            ELSIF (M1Position_M >= (ControlStartM1Position_M + ControlAscentDistance_M))
               AND (M2Position_M >= (ControlStartM2Position_M + ControlAscentDistance_M)) THEN
                ExtractionState := E_ExtractionSequenceState.NOMINAL_ASCENT;
            END_IF;

        E_ExtractionSequenceState.NOMINAL_ASCENT:
            Status.State := E_State.BUSY;
            Status.Busy := TRUE;
            AscentPermit := MotionRequestActive AND (MotionDirection = 1);
            OperatorActionId := 16#0204;
            OperatorAction := 'Maintenir la montée : extraction en cours.';
            IF WinchSyncError OR NOT PositionsValid THEN
                Status.ErrorId := Status.ErrorId OR 16#0004;
                Status.StateAtError := Status.State;
            END_IF;

        E_ExtractionSequenceState.ERROR_HOLD:
            Status.State := E_State.READY;
    END_CASE;
END_IF;

Status.Error := (Status.ErrorId <> 16#0000);

{endregion}
